Staubli VAL3: CheckTraj.pgx

program CheckTraj(point x_pStart, trsf x_trOffset, point x_pEnd, bool& x_bTrajOK)
  local bool l_bOk
  local bool l_bOut
  local num l_nStep
  local trsf l_trMiniOffset
  local trsf l_trStepOffset
  local num l_nVal
  local point l_pTarget
  local jointRs l_jNearBy
  local jointRs l_jTarget
  local jointRs l_jStart
  local point l_pNearBy
  local string l_sPopMsg
begin
  l_trMiniOffset={x_trOffset.x/1000,x_trOffset.y/1000,x_trOffset.z/1000,x_trOffset.rx/1000,x_trOffset.ry/1000,x_trOffset.rz/1000}
  x_pEnd=appro(x_pStart,x_trOffset)
  l_nStep=0
  l_nVal=1
  do
    switch l_nStep
      //******************************************************************
      //Check NearBy Position
      case 0
        l_bOk=pointToJoint(utCurrentTool.tValue,herej(),x_pStart,l_jStart)
        if l_bOk==true
          l_nStep=1
        else
          l_nStep=99
        endIf
      break
      //
      case 1
        l_pNearBy=appro(x_pStart,l_trMiniOffset)
        l_bOk=pointToJoint(utCurrentTool.tValue,herej(),l_pNearBy,l_jNearBy)
        if l_bOk==true
          l_nStep=2
        else
          l_nStep=99
        endIf
      break
      //******************************************************************
      //******************************************************************
      case 2
        l_trStepOffset={x_trOffset.x*l_nVal/100,x_trOffset.y*l_nVal/100,x_trOffset.z*l_nVal/100,x_trOffset.rx*l_nVal/100,x_trOffset.ry*l_nVal/100,x_trOffset.rz*l_nVal/100}
        l_pTarget=appro(x_pStart,l_trStepOffset)
        l_bOk=pointToJoint(utCurrentTool.tValue,herej(),l_pTarget,l_jTarget)
        if l_bOk==true
          l_nStep=3
        else
          l_nStep=99
        endIf
      break
      //
      case 3
        if l_jNearBy.j4-l_jStart.j4>=0 and l_jTarget.j4-l_jStart.j4<0
          l_jTarget.j4=l_jTarget.j4+360
        endIf
        if l_jNearBy.j4-l_jStart.j4<0 and l_jTarget.j4-l_jStart.j4>=0
          l_jTarget.j4=l_jTarget.j4-360
        endIf
        l_nStep=4
      break
      //
      case 4
        if isInRange(l_jTarget)==true
          l_nStep=5
        else
          l_nStep=99
        endIf
      break
      //
      case 5
        if l_nVal<100
          l_nVal=l_nVal+1
          l_nStep=2
        else
          l_nStep=100
        endIf
      break
      //******************************************************************
      case 99
        call updateStr(121,l_sPopMsg,"The maximum rotation angle is only:")
        l_nVal=l_nVal-1
        l_sPopMsg=l_sPopMsg+toString(".",roundDown(l_nVal))+"°"
        popUpMsg(l_sPopMsg)
        //
        x_bTrajOK=false
        l_bOut=true
      break
      case 100
        x_bTrajOK=true
        l_bOut=true
      break
    endSwitch
  until l_bOut
end
